// TIA Portal V21 export
DATA_BLOCK "PosControl_horizontale Achse"   // DB3
// stored: InstanceOfName BasicPosControl, OfSystemLibElement BasicPosControl, OfSystemLibVersion 2.1
BasicPosControl   // technology object, version 2.1
   // VAR_INPUT
   //    ModePos : Int;
   //    EnableAxis : Bool;
   //    CancelTraversing : Bool;
   //    IntermediateStop : Bool;
   //    Positive : Bool;
   //    Negative : Bool;
   //    Jog1 : Bool;
   //    Jog2 : Bool;
   //    FlyRef : Bool;
   //    AckError : Bool;
   //    ExecuteMode : Bool;
   //    Position : LReal;
   //    Velocity : LReal;
   //    OverV : Int;
   //    OverAcc : Int;
   //    OverDec : Int;
   //    ConfigEPos : DWord := 16#0000_000F;
   //    UserSetPZD : Word;
   // END_VAR
   // VAR_OUTPUT
   //    AxisEnabled : Bool;
   //    AxisPosOk : Bool;
   //    AxisSpFixed : Bool;
   //    AxisRef : Bool;
   //    AxisWarn : Bool;
   //    AxisError : Bool;
   //    Lockout : Bool;
   //    ActVelocity : LReal;
   //    ActPosition : LReal;
   //    ActMode : Int;
   //    EPosZSW1 : Word;
   //    EPosZSW2 : Word;
   //    ActWarn : Word;
   //    ActFault : Word;
   //    Error : Bool;
   //    Status : Word;
   //    DiagID : Word;
   //    UserReceivePZD : Word;
   // END_VAR
   // VAR
   //    sbOff1Edge : Bool;
   //    sbOff1 : Bool;
   //    sbExecuteEdge : Bool;
   //    sbExecute : Bool;
   //    sbRefTypEdge : Bool;
   //    sbRefTyp : Bool;
   //    sbMdiStart : Bool;
   //    sbMdiStartEdge : Bool;
   //    sbRefStart : Bool;
   //    sbJogInc : Bool;
   //    sbReady : Bool;
   //    sbIOp : Bool;
   //    sbAccel : Bool;
   //    sbDecel : Bool;
   //    sbAlarm : Bool;
   //    sbFault : Bool;
   //    sbFWD : Bool;
   //    sbBWD : Bool;
   //    sbBusy : Bool;
   //    swStatus : Word;
   //    swEPosZSW1 : Word;
   //    swEPosZSW2 : Word := 16#0000;
   //    siExecuteCyc : Int;
   //    siRefTypCyc : Int;
   //    siJogIncCyc : Int;
   //    siMdiStartCyc : Int;
   //    siRefActRetry : Int;
   //    siModePos : Int;
   //    siModePosMax : Int;
   //    siCycWait : Int;
   //    siRetryMax : Int;
   //    sbModePos : Bool;
   //    STW1 : Word;
   //    EPosSTW1 : Word;
   //    EPosSTW2 : Word := WORD#16#C200;
   //    STW2 : Word;
   //    OverrideV : Word;
   //    PositionSP : DWord;
   //    VelocitySP : DWord;
   //    OverrideA : Word;
   //    OverrideD : Word;
   //    SendPZD12 : Word;
   //    ZSW1 : Word;
   //    EPosZSW3 : Word;
   //    EPosZSW4 : Word;
   //    ZSW2 : Word;
   //    NotUsed : Word;
   //    PositionAV : DWord;
   //    VelocityAV : DWord;
   //    ErrNr : Word;
   //    WarnNr : Word;
   //    ReceivePZD12 : Word;
   //    HWIDSTW : HW_IO := 273;
   //    HWIDZSW : HW_IO := 273;
   //    srResolutionFactor : LReal := 20000.0;
   //    srVelocityFactor : LReal := 1200.0;
   //    srNIST_BFactor : LReal := 0.000111758708953857;
   // END_VAR
BEGIN
END_DATA_BLOCK
